(* IEC 61131-3 sources: llm-plc-st-eval/data/definitivo/qwen2.5-coder_14b/I6/few_shot, 3 files *)

(* ---- ejec_1.st ---- *)
FUNCTION_BLOCK FB_Temperatura
VAR_INPUT
    rawTemp : INT; (* Valor de temperatura crudo *)
END_VAR
VAR_OUTPUT
    tempC : REAL; (* Temperatura en Celsius *)
    enfriador : BOOL; (* Estado del enfriador *)
    almSensor : BOOL; (* Alarma del sensor *)
END_VAR
VAR
    tempMin : REAL := 0.0; (* Temperatura mínima *)
    tempMax : REAL := 100.0; (* Temperatura máxima *)
    rawTempMin : INT := 0; (* Valor mínimo de rawTemp *)
    rawTempMax : INT := 27648; (* Valor máximo de rawTemp *)
    histeresis : REAL := 5.0; (* Histéresis *)
END_VAR

(* Calcula la temperatura en Celsius *)
tempC := (rawTemp - rawTempMin) * (tempMax - tempMin) / (rawTempMax - rawTempMin) + tempMin;

(* Alarma del sensor si rawTemp está fuera de rango *)
almSensor := (rawTemp < rawTempMin) OR (rawTemp > rawTempMax);

(* Control del enfriador con histéresis *)
IF tempC >= 80.0 THEN
    enfriador := TRUE;
ELSIF tempC <= 75.0 THEN
    enfriador := FALSE;
END_IF;
END_FUNCTION_BLOCK

(* ---- ejec_2.st ---- *)
FUNCTION_BLOCK FB_Temperatura
VAR_INPUT
    rawTemp : INT; (* Valor raw de temperatura *)
END_VAR
VAR_OUTPUT
    tempC : REAL; (* Temperatura en Celsius *)
    enfriador : BOOL; (* Control del enfriador *)
    almSensor : BOOL; (* Alarma del sensor *)
END_VAR
VAR
    tempMin : REAL := 0.0; (* Temperatura mínima *)
    tempMax : REAL := 100.0; (* Temperatura máxima *)
    rawMin : INT := 0; (* Valor raw mínimo *)
    rawMax : INT := 27648; (* Valor raw máximo *)
    tempThresholdHigh : REAL := 80.0; (* Umbral alto para activar el enfriador *)
    tempThresholdLow : REAL := 75.0; (* Umbral bajo para desactivar el enfriador *)
END_VAR

(* Conversión de rawTemp a temperatura en Celsius *)
tempC := (rawTemp - rawMin) * (tempMax - tempMin) / (rawMax - rawMin) + tempMin;

(* Control del enfriador con histéresis *)
IF tempC >= tempThresholdHigh THEN
    enfriador := TRUE;
ELSIF tempC <= tempThresholdLow THEN
    enfriador := FALSE;
END_IF;

(* Alarma del sensor si rawTemp está fuera de rango *)
IF rawTemp < rawMin OR rawTemp > rawMax THEN
    almSensor := TRUE;
    enfriador := FALSE;
ELSE
    almSensor := FALSE;
END_IF;
END_FUNCTION_BLOCK

(* ---- ejec_3.st ---- *)
FUNCTION_BLOCK FB_Temperatura
VAR_INPUT
    rawTemp : INT; (* Valor raw de temperatura *)
END_VAR
VAR_OUTPUT
    tempC : REAL; (* Temperatura en grados Celsius *)
    enfriador : BOOL; (* Estado del enfriador *)
    almSensor : BOOL; (* Alarma de sensor *)
END_VAR
VAR
    tempMin : REAL := 0.0; (* Temperatura mínima *)
    tempMax : REAL := 100.0; (* Temperatura máxima *)
    rawMin : INT := 0; (* Valor raw mínimo *)
    rawMax : INT := 27648; (* Valor raw máximo *)
    tempThresholdHigh : REAL := 80.0; (* Umbral alto para activar el enfriador *)
    tempThresholdLow : REAL := 75.0; (* Umbral bajo para desactivar el enfriador *)
END_VAR

(* Conversión de rawTemp a temperatura en Celsius *)
IF rawTemp < rawMin OR rawTemp > rawMax THEN
    almSensor := TRUE;
    tempC := 0.0;
    enfriador := FALSE;
ELSE
    almSensor := FALSE;
    tempC := (rawTemp - rawMin) * (tempMax - tempMin) / (rawMax - rawMin) + tempMin;
    (* Control del enfriador con histéresis *)
    IF tempC >= tempThresholdHigh THEN
        enfriador := TRUE;
    ELSIF tempC <= tempThresholdLow THEN
        enfriador := FALSE;
    END_IF;
END_IF;
END_FUNCTION_BLOCK
